Fanuc KAREL source: KA00194.KL

PROGRAM KA00194
%NOLOCKGROUP
VAR
  SRC: ARRAY[4] OF SHORT
  DST: ARRAY[4] OF BYTE
BEGIN
  DST = SRC
END KA00194
